// TIA Portal V20 export
// export: Created 2026-10-20T12:44:48.0111089Z, ExportSetting WithDefaults, DisplayName Totally Integrated Automation Portal, DisplayVersion V20 Update 6, DisplayName TIA Portal Openness, DisplayVersion V20 Update 6, DisplayName TIA Portal Version Control Interface, DisplayVersion V20 Update 6, DisplayName SINAMICS Startdrive Advanced, DisplayVersion V20 SP1, DisplayName SINAMICS Startdrive G130, G150, S120, S150, SINAMICS MV, G220, S200, S210, DisplayVersion V20 SP1, DisplayName SINAMICS Startdrive G110M, G120, G120C, G120D, G120P, G115D, DisplayVersion V20 SP1, DisplayName STEP 7 Professional, DisplayVersion V20 Update 6, DisplayName STEP 7 Safety, DisplayVersion V20 Update 2, DisplayName WinCC Basic/Comfort/Advanced, DisplayVersion V20 Update 6, DisplayName WinCC Unified, DisplayVersion V20 Update 6
FUNCTION "OT_Charge_Commands_1" : Void   // FC64, SCL
{ S7_Optimized_Access := 'TRUE' }
VERSION : 0.1
// stored: AutoNumber true, IsIECCheckEnabled false, SetENOAutomatically false, UDAEnableTagReadback false
   VAR_IN_OUT
      Auto_Test : "Auto_Test_1";
   END_VAR
BEGIN
   "OrderTable_HMI"."Manual order" := #Auto_Test.Manual;
   //PALLET TYPE
   IF #Auto_Test."Pallet Type" = 'C' THEN
       "OrderTable_HMI"."Pallet Type" := 1;
   ELSIF #Auto_Test."Pallet Type" = 'E' THEN
       "OrderTable_HMI"."Pallet Type" := 2;
   END_IF;
   //TOWER 1 PALLET ALIGNMENT
   IF #Auto_Test."Tower 1 Pallet Alignment" = 'R' THEN
       "OrderTable_HMI"."Tower 1 Pallet Alignment" := 1;
   ELSIF #Auto_Test."Tower 1 Pallet Alignment" = 'L' THEN
       "OrderTable_HMI"."Tower 1 Pallet Alignment" := 2;
   END_IF;
   //ECONVEYOR PALLET ALIGNMENT
   IF #Auto_Test."Extractor Pallet Alignment" = 'R' THEN
       "OrderTable_HMI"."Extractor Pallet Alignment" := 1;
   ELSIF #Auto_Test."Extractor Pallet Alignment" = 'L' THEN
       "OrderTable_HMI"."Extractor Pallet Alignment" := 2;
   ELSIF #Auto_Test."Extractor Pallet Alignment" = 'C' THEN
       "OrderTable_HMI"."Extractor Pallet Alignment" := 3;
   END_IF;
   "OrderTable_HMI"."From level" := #Auto_Test."From level";
   "OrderTable_HMI"."To level" := #Auto_Test."To level";
   "OrderTable_HMI"."Testing Time" := #Auto_Test."Testing Time";
   "OrderTable_HMI"."Numer of cycles" := #Auto_Test."Numer of cycles";
   "OrderTable_HMI".Level := UINT_TO_BYTE(#Auto_Test.Level);
   "OrderTable_HMI".Tower := UINT_TO_BYTE(#Auto_Test.Tower);
END_FUNCTION
